(* IEC 61131-3 sources: avi-aoi-management/scripts/ai-eval/ngau-nhien/kho/st-ud1-bom-luan-phien/khung/src, 2 files *)

(* ---- BomLuanPhien.st ---- *)
FUNCTION_BLOCK BomLuanPhien
VAR_INPUT
    MUC_CAO : BOOL;
    MUC_THAP : BOOL;
    PH1 : BOOL;
    PH2 : BOOL;
    RESET : BOOL;
    T_PHAN_HOI : TIME;
END_VAR
VAR_OUTPUT
    BOM1 : BOOL;
    BOM2 : BOOL;
    CAN_BOM : BOOL;
    LOI1 : BOOL;
    LOI2 : BOOL;
    BAO_DONG : BOOL;
    BOM_CHINH : INT;
END_VAR
    (* TODO: cài đặt theo đề bài *)
    BOM1 := FALSE;
END_FUNCTION_BLOCK

(* ---- GiamSatBom.st ---- *)
FUNCTION_BLOCK GiamSatBom
VAR_INPUT
    LENH : BOOL;
    PHAN_HOI : BOOL;
    RESET : BOOL;
    T_PHAN_HOI : TIME;
END_VAR
VAR_OUTPUT
    LOI : BOOL;
END_VAR
    (* TODO: cài đặt theo đề bài *)
    LOI := FALSE;
END_FUNCTION_BLOCK
